// TIA Portal V20 export
DATA_BLOCK "Verwaltung_Teiledaten"   // DB2
{ S7_Optimized_Access := 'TRUE' }
// stored: MemoryReserve 100
   VAR RETAIN
      Artikel_gewechselt : Bool;
      Datensatz : String;
      Rezeptnummer : String;
      "Achse Position GS" : Real;   // Achse Position GS [mm]
      "Achse Position AS" : Real;   // Achse Position GS [mm]
      "Achse Geschwindigkeit GS->AS" : Real;   // Achse Geschwindigkeit GS->AS [mm/min]
      "Achse Geschwindigkeit AS->GS" : Real;   // Achse Geschwindigkeit AS->GS [mm/min]
      "Drehantrieb Position GS" : Real;   // Drehantrieb Position GS [°]
      "Drehantrieb Position AS1" : Real;   // Drehantrieb Position AS1 [°]
      "Drehantrieb Position AS2" : Real;   // Drehantrieb Position AS1 [°]
      "Drehantrieb Geschwindigkeit GS->AS1" : Real;   // Drehantrieb Geschwindigkeit GS->AS1 [°/s]
      "Drehantrieb Geschwindigkeit AS1->GS" : Real;   // Drehantrieb Geschwindigkeit AS1->GS [°/s]
      "Wartezeit gesteckt" : Real;   // Wartezeit gesteckt [s]
      "Drehantrieb Motorstrombegrenzung" : Real;   // Drehantrieb Motorstrombegrenzung [%]
      "Druck p1 Ausgleichszylinder" : Int;   // Druck p1 Ausgleichszylinder [bar]
      "Druck p2 Überlastzylinder" : Int;   // Druck p2 Überlastzylinder [bar]
      "Wegmessung_Ausgleichszylinder Position GS" : Real;   // Wegmessung Ausgleichszylinder Position GS [mm]
      "Wegmessung_Ausgleichszylinder Position AS1" : Real;   // Wegmessung Ausgleichszylinder Position AS1 [mm]
      "Wegmessung_Ausgleichszylinder maximale Abweichung GS" : Real;   // Wegmessung Ausgleichszylinder maximale Abweichung GS [mm]
      "Wegmessung_Ausgleichszylinder maximale Abweichung AS1" : Real;   // Wegmessung Ausgleichszylinder maximale Abweichung AS1 [mm]
      "Taster Achse Position GS übernehmen" : Bool;   // Taster Achse Position GS übernehmen
      "Taster Achse Position AS übernehmen" : Bool;   // Taster Achse Position AS übernehmen
      "Taster Drehantrieb Position GS übernehmen" : Bool;   // Taster Drehantrieb Position GS übernehmen
      "Taster Drehantrieb Position AS1 übernehmen" : Bool;   // Taster Drehantrieb Position AS1 übernehmen
      "Taster Drehantrieb Position AS2 übernehmen" : Bool;   // Taster Drehantrieb Position AS2 übernehmen
      "Taster Wegmessung Ausgleichszylinder Position GS übernehmen" : Bool;   // Taster Wegmessung Ausgleichszylinder Position GS übernehmen
      "Taster Wegmessung Ausgleichszylinder Position AS1 übernehmen" : Bool;   // Taster Wegmessung Ausgleichszylinder Position AS1 übernehmen
   END_VAR
BEGIN
END_DATA_BLOCK
